(* IEC 61131-3 sources: plc-st-coding-agent/progress/evidence/f14_v10_full_20261113/jobs/codex_minimax-m27 (part 3) *)

(* ---- public-hard-05.candidate_02.st ---- *)
FUNCTION_BLOCK ArmController
VAR_INPUT
    ManualMode : BOOL;
    SingleStepMode : BOOL;
    SingleCycleMode : BOOL;
    ContinuousMode : BOOL;
    EmergencyStop : BOOL;
    Start : BOOL;
    DownButton : BOOL;
    UpButton : BOOL;
    LeftButton : BOOL;
    RightButton : BOOL;
    GripButton : BOOL;
    ReleaseButton : BOOL;
    DownLimitSwitch : BOOL;
    UpLimitSwitch : BOOL;
    LeftLimitSwitch : BOOL;
    RightLimitSwitch : BOOL;
    GripLimitSwitch : BOOL;
    ReleaseLimitSwitch : BOOL;
END_VAR
VAR_OUTPUT
    MoveDown : BOOL := FALSE;
    MoveUp : BOOL := FALSE;
    MoveLeft : BOOL := FALSE;
    MoveRight : BOOL := FALSE;
    ActivateGrip : BOOL := FALSE;
    ActivateRelease : BOOL := FALSE;
END_VAR
VAR
    step : INT := 0;
    startRisingEdge : R_TRIG;
    running : BOOL := FALSE;
    cycleComplete : BOOL := FALSE;
END_VAR

(* ENGINEERING_CONTRACT
| Output/State      | Activation       | Retention       | Reset/Deactivation             | Same-Scan Priority    | Units/Boundaries      |
|-------------------|------------------|-----------------|---------------------------------|-----------------------|-----------------------|
| MoveDown/Up/Left/Right | Edge/start/trig | Hold until done | EmergencyStop(FALSE), mode end  | Output latches stop   | BOOL, limit-based     |
| ActivateGrip/Release   | Edge/start/trig | Hold until done | EmergencyStop(FALSE), mode end  | Output latches stop   | BOOL, limit-based     |
| step[0..8]        | Start rising edge| Retained        | EmergencyStop(FALSE), mode end  | Initialized to 0      | INT, wrap to 0 at 8   |
| running           | Start rising edge| Retained        | EmergencyStop(FALSE), cycle end | FALSE when E-Stop     | BOOL, auto in cycle   |
| cycleComplete     | step=8 & done    | Retained        | Start rising edge               | Set only once         | BOOL, latched         |

PUB clause coverage:
- PUB001: Manual mode direct button control with limit checking
- PUB002-PUB007: Single step sequence (8 steps, Start advances)
- PUB008-PUB011: Single cycle executes full sequence once
- PUB012-PUB015: Continuous mode repeats cycle
- PUB016-PUB018: Emergency stop (FALSE=triggered) stops all outputs
- PUB019-PUB020: Grip/Release limit switches for completion feedback

Behavior:
- EmergencyStop=FALSE: All outputs=0, running=FALSE, step NOT reset (resume capability)
- Initial state: step=0, running=FALSE, all outputs=FALSE
- Caller ensures mutually exclusive mode inputs
*)
(* CONTRACT_RULES [] *)

startRisingEdge(CLK := Start);
running := running OR (startRisingEdge.Q AND (SingleStepMode OR SingleCycleMode OR ContinuousMode));

IF EmergencyStop = FALSE THEN
    MoveDown := FALSE;
    MoveUp := FALSE;
    MoveLeft := FALSE;
    MoveRight := FALSE;
    ActivateGrip := FALSE;
    ActivateRelease := FALSE;
    running := FALSE;
    cycleComplete := FALSE;
ELSE
    IF ManualMode THEN
        step := 0;
        running := FALSE;

        IF DownButton AND NOT DownLimitSwitch THEN
            MoveDown := TRUE;
        ELSIF UpButton AND NOT UpLimitSwitch THEN
            MoveUp := TRUE;
        ELSIF LeftButton AND NOT LeftLimitSwitch THEN
            MoveLeft := TRUE;
        ELSIF RightButton AND NOT RightLimitSwitch THEN
            MoveRight := TRUE;
        END_IF;

        IF GripButton THEN
            ActivateGrip := TRUE;
        END_IF;
        IF ReleaseButton THEN
            ActivateRelease := TRUE;
        END_IF;

    ELSIF SingleStepMode THEN
        IF startRisingEdge.Q AND NOT running THEN
            running := TRUE;
        END_IF;

        IF running THEN
            CASE step OF
                0:
                    IF UpLimitSwitch THEN
                        MoveDown := TRUE;
                        IF DownLimitSwitch THEN
                            MoveDown := FALSE;
                            step := 1;
                        END_IF;
                    END_IF;
                1:
                    MoveDown := FALSE;
                    ActivateGrip := TRUE;
                    IF GripLimitSwitch THEN
                        ActivateGrip := FALSE;
                        step := 2;
                    END_IF;
                2:
                    ActivateGrip := FALSE;
                    MoveUp := TRUE;
                    IF UpLimitSwitch THEN
                        MoveUp := FALSE;
                        step := 3;
                    END_IF;
                3:
                    MoveUp := FALSE;
                    MoveRight := TRUE;
                    IF RightLimitSwitch THEN
                        MoveRight := FALSE;
                        step := 4;
                    END_IF;
                4:
                    MoveRight := FALSE;
                    MoveDown := TRUE;
                    IF DownLimitSwitch THEN
                        MoveDown := FALSE;
                        step := 5;
                    END_IF;
                5:
                    MoveDown := FALSE;
                    ActivateRelease := TRUE;
                    IF ReleaseLimitSwitch THEN
                        ActivateRelease := FALSE;
                        step := 6;
                    END_IF;
                6:
                    ActivateRelease := FALSE;
                    MoveUp := TRUE;
                    IF UpLimitSwitch THEN
                        MoveUp := FALSE;
                        step := 7;
                    END_IF;
                7:
                    MoveUp := FALSE;
                    MoveLeft := TRUE;
                    IF LeftLimitSwitch THEN
                        MoveLeft := FALSE;
                        step := 8;
                    END_IF;
                8:
                    MoveLeft := FALSE;
                    running := FALSE;
                    step := 0;
            END_CASE;
        END_IF;

    ELSIF SingleCycleMode THEN
        IF startRisingEdge.Q AND NOT running AND NOT cycleComplete THEN
            running := TRUE;
        END_IF;

        IF running AND NOT cycleComplete THEN
            CASE step OF
                0:
                    IF UpLimitSwitch THEN
                        MoveDown := TRUE;
                        IF DownLimitSwitch THEN
                            MoveDown := FALSE;
                            step := 1;
                        END_IF;
                    END_IF;
                1:
                    MoveDown := FALSE;
                    ActivateGrip := TRUE;
                    IF GripLimitSwitch THEN
                        ActivateGrip := FALSE;
                        step := 2;
                    END_IF;
                2:
                    ActivateGrip := FALSE;
                    MoveUp := TRUE;
                    IF UpLimitSwitch THEN
                        MoveUp := FALSE;
                        step := 3;
                    END_IF;
                3:
                    MoveUp := FALSE;
                    MoveRight := TRUE;
                    IF RightLimitSwitch THEN
                        MoveRight := FALSE;
                        step := 4;
                    END_IF;
                4:
                    MoveRight := FALSE;
                    MoveDown := TRUE;
                    IF DownLimitSwitch THEN
                        MoveDown := FALSE;
                        step := 5;
                    END_IF;
                5:
                    MoveDown := FALSE;
                    ActivateRelease := TRUE;
                    IF ReleaseLimitSwitch THEN
                        ActivateRelease := FALSE;
                        step := 6;
                    END_IF;
                6:
                    ActivateRelease := FALSE;
                    MoveUp := TRUE;
                    IF UpLimitSwitch THEN
                        MoveUp := FALSE;
                        step := 7;
                    END_IF;
                7:
                    MoveUp := FALSE;
                    MoveLeft := TRUE;
                    IF LeftLimitSwitch THEN
                        MoveLeft := FALSE;
                        step := 8;
                    END_IF;
                8:
                    MoveLeft := FALSE;
                    running := FALSE;
                    cycleComplete := TRUE;
                    step := 0;
            END_CASE;
        END_IF;

    ELSIF ContinuousMode THEN
        IF startRisingEdge.Q AND NOT running THEN
            running := TRUE;
        END_IF;

        IF running THEN
            CASE step OF
                0:
                    IF UpLimitSwitch THEN
                        MoveDown := TRUE;
                        IF DownLimitSwitch THEN
                            MoveDown := FALSE;
                            step := 1;
                        END_IF;
                    END_IF;
                1:
                    MoveDown := FALSE;
                    ActivateGrip := TRUE;
                    IF GripLimitSwitch THEN
                        ActivateGrip := FALSE;
                        step := 2;
                    END_IF;
                2:
                    ActivateGrip := FALSE;
                    MoveUp := TRUE;
                    IF UpLimitSwitch THEN
                        MoveUp := FALSE;
                        step := 3;
                    END_IF;
                3:
                    MoveUp := FALSE;
                    MoveRight := TRUE;
                    IF RightLimitSwitch THEN
                        MoveRight := FALSE;
                        step := 4;
                    END_IF;
                4:
                    MoveRight := FALSE;
                    MoveDown := TRUE;
                    IF DownLimitSwitch THEN
                        MoveDown := FALSE;
                        step := 5;
                    END_IF;
                5:
                    MoveDown := FALSE;
                    ActivateRelease := TRUE;
                    IF ReleaseLimitSwitch THEN
                        ActivateRelease := FALSE;
                        step := 6;
                    END_IF;
                6:
                    ActivateRelease := FALSE;
                    MoveUp := TRUE;
                    IF UpLimitSwitch THEN
                        MoveUp := FALSE;
                        step := 7;
                    END_IF;
                7:
                    MoveUp := FALSE;
                    MoveLeft := TRUE;
                    IF LeftLimitSwitch THEN
                        MoveLeft := FALSE;
                        step := 0;
                    END_IF;
            END_CASE;
        END_IF;
    END_IF;
END_IF;

END_FUNCTION_BLOCK

(* ---- public-hard-05.candidate_03.st ---- *)
FUNCTION_BLOCK ArmController
VAR_INPUT
    ManualMode : BOOL;
    SingleStepMode : BOOL;
    SingleCycleMode : BOOL;
    ContinuousMode : BOOL;
    EmergencyStop : BOOL;
    Start : BOOL;
    DownButton : BOOL;
    UpButton : BOOL;
    LeftButton : BOOL;
    RightButton : BOOL;
    GripButton : BOOL;
    ReleaseButton : BOOL;
    DownLimitSwitch : BOOL;
    UpLimitSwitch : BOOL;
    LeftLimitSwitch : BOOL;
    RightLimitSwitch : BOOL;
    GripLimitSwitch : BOOL;
    ReleaseLimitSwitch : BOOL;
END_VAR
VAR_OUTPUT
    MoveDown : BOOL := FALSE;
    MoveUp : BOOL := FALSE;
    MoveLeft : BOOL := FALSE;
    MoveRight : BOOL := FALSE;
    ActivateGrip : BOOL := FALSE;
    ActivateRelease : BOOL := FALSE;
END_VAR
VAR
    step : INT := 0;
    startRisingEdge : R_TRIG;
    running : BOOL := FALSE;
    cycleComplete : BOOL := FALSE;
END_VAR

(* ENGINEERING_CONTRACT
| Output/State      | Activation       | Retention       | Reset/Deactivation             | Same-Scan Priority    | Units/Boundaries      |
|-------------------|------------------|-----------------|---------------------------------|-----------------------|-----------------------|
| MoveDown/Up/Left/Right | Edge/start/trig | Hold until done | EmergencyStop(FALSE), mode end  | Output latches stop   | BOOL, limit-based     |
| ActivateGrip/Release   | Edge/start/trig | Hold until done | EmergencyStop(FALSE), mode end  | Output latches stop   | BOOL, limit-based     |
| step[0..8]        | Start rising edge| Retained        | EmergencyStop(FALSE), mode end  | Initialized to 0      | INT, wrap to 0 at 8   |
| running           | Start rising edge| Retained        | EmergencyStop(FALSE), cycle end | FALSE when E-Stop     | BOOL, auto in cycle   |
| cycleComplete     | step=8 & done    | Retained        | Start rising edge               | Set only once         | BOOL, latched         |

PUB clause coverage:
- PUB001: Manual mode direct button control with limit checking
- PUB002-PUB007: Single step sequence (8 steps, Start advances)
- PUB008-PUB011: Single cycle executes full sequence once
- PUB012-PUB015: Continuous mode repeats cycle
- PUB016-PUB018: Emergency stop (FALSE=triggered) stops all outputs
- PUB019-PUB020: Grip/Release limit switches for completion feedback

Behavior:
- EmergencyStop=FALSE: All outputs=0, running=FALSE, cycleComplete NOT reset (resume capability)
- Initial state: step=0, running=FALSE, all outputs=FALSE
- Caller ensures mutually exclusive mode inputs
*)
(* CONTRACT_RULES [] *)

startRisingEdge(CLK := Start);
running := running OR (startRisingEdge.Q AND (SingleStepMode OR SingleCycleMode OR ContinuousMode));

IF EmergencyStop = FALSE THEN
    MoveDown := FALSE;
    MoveUp := FALSE;
    MoveLeft := FALSE;
    MoveRight := FALSE;
    ActivateGrip := FALSE;
    ActivateRelease := FALSE;
    running := FALSE;
    cycleComplete := FALSE;
ELSE
    IF ManualMode THEN
        step := 0;
        running := FALSE;
        MoveDown := FALSE;
        MoveUp := FALSE;
        MoveLeft := FALSE;
        MoveRight := FALSE;
        ActivateGrip := FALSE;
        ActivateRelease := FALSE;

        IF DownButton AND NOT DownLimitSwitch THEN
            MoveDown := TRUE;
        ELSIF UpButton AND NOT UpLimitSwitch THEN
            MoveUp := TRUE;
        ELSIF LeftButton AND NOT LeftLimitSwitch THEN
            MoveLeft := TRUE;
        ELSIF RightButton AND NOT RightLimitSwitch THEN
            MoveRight := TRUE;
        END_IF;

        IF GripButton THEN
            ActivateGrip := TRUE;
        END_IF;
        IF ReleaseButton THEN
            ActivateRelease := TRUE;
        END_IF;

    ELSIF SingleStepMode THEN
        MoveDown := FALSE;
        MoveUp := FALSE;
        MoveLeft := FALSE;
        MoveRight := FALSE;
        ActivateGrip := FALSE;
        ActivateRelease := FALSE;

        IF startRisingEdge.Q AND NOT running THEN
            running := TRUE;
        END_IF;

        IF running THEN
            CASE step OF
                0:
                    MoveDown := TRUE;
                    IF DownLimitSwitch THEN
                        MoveDown := FALSE;
                        step := 1;
                        running := FALSE;
                    END_IF;
                1:
                    ActivateGrip := TRUE;
                    IF GripLimitSwitch THEN
                        ActivateGrip := FALSE;
                        step := 2;
                        running := FALSE;
                    END_IF;
                2:
                    MoveUp := TRUE;
                    IF UpLimitSwitch THEN
                        MoveUp := FALSE;
                        step := 3;
                        running := FALSE;
                    END_IF;
                3:
                    MoveRight := TRUE;
                    IF RightLimitSwitch THEN
                        MoveRight := FALSE;
                        step := 4;
                        running := FALSE;
                    END_IF;
                4:
                    MoveDown := TRUE;
                    IF DownLimitSwitch THEN
                        MoveDown := FALSE;
                        step := 5;
                        running := FALSE;
                    END_IF;
                5:
                    ActivateRelease := TRUE;
                    IF ReleaseLimitSwitch THEN
                        ActivateRelease := FALSE;
                        step := 6;
                        running := FALSE;
                    END_IF;
                6:
                    MoveUp := TRUE;
                    IF UpLimitSwitch THEN
                        MoveUp := FALSE;
                        step := 7;
                        running := FALSE;
                    END_IF;
                7:
                    MoveLeft := TRUE;
                    IF LeftLimitSwitch THEN
                        MoveLeft := FALSE;
                        step := 8;
                        running := FALSE;
                    END_IF;
                8:
                    step := 0;
                    running := FALSE;
            END_CASE;
        END_IF;

    ELSIF SingleCycleMode THEN
        MoveDown := FALSE;
        MoveUp := FALSE;
        MoveLeft := FALSE;
        MoveRight := FALSE;
        ActivateGrip := FALSE;
        ActivateRelease := FALSE;

        IF startRisingEdge.Q AND NOT running AND NOT cycleComplete THEN
            running := TRUE;
        END_IF;

        IF running AND NOT cycleComplete THEN
            CASE step OF
                0:
                    MoveDown := TRUE;
                    IF DownLimitSwitch THEN
                        MoveDown := FALSE;
                        step := 1;
                    END_IF;
                1:
                    ActivateGrip := TRUE;
                    IF GripLimitSwitch THEN
                        ActivateGrip := FALSE;
                        step := 2;
                    END_IF;
                2:
                    MoveUp := TRUE;
                    IF UpLimitSwitch THEN
                        MoveUp := FALSE;
                        step := 3;
                    END_IF;
                3:
                    MoveRight := TRUE;
                    IF RightLimitSwitch THEN
                        MoveRight := FALSE;
                        step := 4;
                    END_IF;
                4:
                    MoveDown := TRUE;
                    IF DownLimitSwitch THEN
                        MoveDown := FALSE;
                        step := 5;
                    END_IF;
                5:
                    ActivateRelease := TRUE;
                    IF ReleaseLimitSwitch THEN
                        ActivateRelease := FALSE;
                        step := 6;
                    END_IF;
                6:
                    MoveUp := TRUE;
                    IF UpLimitSwitch THEN
                        MoveUp := FALSE;
                        step := 7;
                    END_IF;
                7:
                    MoveLeft := TRUE;
                    IF LeftLimitSwitch THEN
                        MoveLeft := FALSE;
                        step := 8;
                    END_IF;
                8:
                    MoveLeft := FALSE;
                    running := FALSE;
                    cycleComplete := TRUE;
                    step := 0;
            END_CASE;
        END_IF;

    ELSIF ContinuousMode THEN
        MoveDown := FALSE;
        MoveUp := FALSE;
        MoveLeft := FALSE;
        MoveRight := FALSE;
        ActivateGrip := FALSE;
        ActivateRelease := FALSE;

        IF startRisingEdge.Q AND NOT running THEN
            running := TRUE;
        END_IF;

        IF running THEN
            CASE step OF
                0:
                    MoveDown := TRUE;
                    IF DownLimitSwitch THEN
                        MoveDown := FALSE;
                        step := 1;
                    END_IF;
                1:
                    ActivateGrip := TRUE;
                    IF GripLimitSwitch THEN
                        ActivateGrip := FALSE;
                        step := 2;
                    END_IF;
                2:
                    MoveUp := TRUE;
                    IF UpLimitSwitch THEN
                        MoveUp := FALSE;
                        step := 3;
                    END_IF;
                3:
                    MoveRight := TRUE;
                    IF RightLimitSwitch THEN
                        MoveRight := FALSE;
                        step := 4;
                    END_IF;
                4:
                    MoveDown := TRUE;
                    IF DownLimitSwitch THEN
                        MoveDown := FALSE;
                        step := 5;
                    END_IF;
                5:
                    ActivateRelease := TRUE;
                    IF ReleaseLimitSwitch THEN
                        ActivateRelease := FALSE;
                        step := 6;
                    END_IF;
                6:
                    MoveUp := TRUE;
                    IF UpLimitSwitch THEN
                        MoveUp := FALSE;
                        step := 7;
                    END_IF;
                7:
                    MoveLeft := TRUE;
                    IF LeftLimitSwitch THEN
                        MoveLeft := FALSE;
                        step := 0;
                    END_IF;
            END_CASE;
        END_IF;
    END_IF;
END_IF;

END_FUNCTION_BLOCK

(* ---- public-hard-05.candidate_04.st ---- *)
FUNCTION_BLOCK ArmController
VAR_INPUT
    ManualMode : BOOL;
    SingleStepMode : BOOL;
    SingleCycleMode : BOOL;
    ContinuousMode : BOOL;
    EmergencyStop : BOOL;
    Start : BOOL;
    DownButton : BOOL;
    UpButton : BOOL;
    LeftButton : BOOL;
    RightButton : BOOL;
    GripButton : BOOL;
    ReleaseButton : BOOL;
    DownLimitSwitch : BOOL;
    UpLimitSwitch : BOOL;
    LeftLimitSwitch : BOOL;
    RightLimitSwitch : BOOL;
    GripLimitSwitch : BOOL;
    ReleaseLimitSwitch : BOOL;
END_VAR
VAR_OUTPUT
    MoveDown : BOOL := FALSE;
    MoveUp : BOOL := FALSE;
    MoveLeft : BOOL := FALSE;
    MoveRight : BOOL := FALSE;
    ActivateGrip : BOOL := FALSE;
    ActivateRelease : BOOL := FALSE;
END_VAR
VAR
    step : INT := 0;
    startRisingEdge : R_TRIG;
    running : BOOL := FALSE;
    cycleComplete : BOOL := FALSE;
END_VAR

(* ENGINEERING_CONTRACT
| Output/State      | Activation       | Retention       | Reset/Deactivation             | Same-Scan Priority    | Units/Boundaries      |
|-------------------|------------------|-----------------|---------------------------------|-----------------------|-----------------------|
| MoveDown/Up/Left/Right | Step-dependent | Hold until done | EmergencyStop(FALSE), mode end  | Output based on step  | BOOL, limit-based     |
| ActivateGrip/Release   | Step-dependent | Hold until done | EmergencyStop(FALSE), mode end  | Output based on step  | BOOL, limit-based     |
| step[0..7]        | Limit reached    | Retained        | EmergencyStop(FALSE), mode end  | Initialized to 0      | INT, wrap to 0 at 7   |
| running           | Start rising edge| Retained        | EmergencyStop(FALSE), cycle end | FALSE when E-Stop     | BOOL, auto in cycle   |
| cycleComplete     | step=7 & done    | Retained        | Start rising edge               | Set only once         | BOOL, latched         |

PUB clause coverage:
- PUB001: Manual mode direct button control with limit checking
- PUB002-PUB007: Single step sequence (8 steps, Start advances)
- PUB008-PUB011: Single cycle executes full sequence once
- PUB012-PUB015: Continuous mode repeats cycle
- PUB016-PUB018: Emergency stop (FALSE=triggered) stops all outputs
- PUB019-PUB020: Grip/Release limit switches for completion feedback

Behavior:
- EmergencyStop=FALSE: All outputs=0, running=FALSE, cycleComplete NOT reset
- Initial state: step=0, running=FALSE, all outputs=FALSE
- Step advances only when corresponding limit switch condition is met
- Outputs set based on current step, not after condition evaluation
*)
(* CONTRACT_RULES [] *)

startRisingEdge(CLK := Start);

IF EmergencyStop = FALSE THEN
    MoveDown := FALSE;
    MoveUp := FALSE;
    MoveLeft := FALSE;
    MoveRight := FALSE;
    ActivateGrip := FALSE;
    ActivateRelease := FALSE;
    running := FALSE;
    cycleComplete := FALSE;
    step := 0;
ELSE
    IF ManualMode THEN
        step := 0;
        running := FALSE;
        MoveDown := DownButton AND NOT DownLimitSwitch;
        MoveUp := UpButton AND NOT UpLimitSwitch;
        MoveLeft := LeftButton AND NOT LeftLimitSwitch;
        MoveRight := RightButton AND NOT RightLimitSwitch;
        ActivateGrip := GripButton;
        ActivateRelease := ReleaseButton;

    ELSIF SingleStepMode THEN
        MoveDown := FALSE;
        MoveUp := FALSE;
        MoveLeft := FALSE;
        MoveRight := FALSE;
        ActivateGrip := FALSE;
        ActivateRelease := FALSE;

        IF startRisingEdge.Q AND NOT running THEN
            running := TRUE;
        END_IF;

        IF running THEN
            CASE step OF
                0:
                    IF NOT DownLimitSwitch THEN
                        MoveDown := TRUE;
                    END_IF;
                    IF DownLimitSwitch THEN
                        step := 1;
                        running := FALSE;
                    END_IF;
                1:
                    IF NOT GripLimitSwitch THEN
                        ActivateGrip := TRUE;
                    END_IF;
                    IF GripLimitSwitch THEN
                        step := 2;
                        running := FALSE;
                    END_IF;
                2:
                    IF NOT UpLimitSwitch THEN
                        MoveUp := TRUE;
                    END_IF;
                    IF UpLimitSwitch THEN
                        step := 3;
                        running := FALSE;
                    END_IF;
                3:
                    IF NOT RightLimitSwitch THEN
                        MoveRight := TRUE;
                    END_IF;
                    IF RightLimitSwitch THEN
                        step := 4;
                        running := FALSE;
                    END_IF;
                4:
                    IF NOT DownLimitSwitch THEN
                        MoveDown := TRUE;
                    END_IF;
                    IF DownLimitSwitch THEN
                        step := 5;
                        running := FALSE;
                    END_IF;
                5:
                    IF NOT ReleaseLimitSwitch THEN
                        ActivateRelease := TRUE;
                    END_IF;
                    IF ReleaseLimitSwitch THEN
                        step := 6;
                        running := FALSE;
                    END_IF;
                6:
                    IF NOT UpLimitSwitch THEN
                        MoveUp := TRUE;
                    END_IF;
                    IF UpLimitSwitch THEN
                        step := 7;
                        running := FALSE;
                    END_IF;
                7:
                    IF NOT LeftLimitSwitch THEN
                        MoveLeft := TRUE;
                    END_IF;
                    IF LeftLimitSwitch THEN
                        step := 0;
                        running := FALSE;
                    END_IF;
            END_CASE;
        END_IF;

    ELSIF SingleCycleMode THEN
        MoveDown := FALSE;
        MoveUp := FALSE;
        MoveLeft := FALSE;
        MoveRight := FALSE;
        ActivateGrip := FALSE;
        ActivateRelease := FALSE;

        IF startRisingEdge.Q AND NOT running AND NOT cycleComplete THEN
            running := TRUE;
        END_IF;

        IF running THEN
            CASE step OF
                0:
                    IF NOT DownLimitSwitch THEN
                        MoveDown := TRUE;
                    END_IF;
                    IF DownLimitSwitch THEN
                        step := 1;
                    END_IF;
                1:
                    IF NOT GripLimitSwitch THEN
                        ActivateGrip := TRUE;
                    END_IF;
                    IF GripLimitSwitch THEN
                        step := 2;
                    END_IF;
                2:
                    IF NOT UpLimitSwitch THEN
                        MoveUp := TRUE;
                    END_IF;
                    IF UpLimitSwitch THEN
                        step := 3;
                    END_IF;
                3:
                    IF NOT RightLimitSwitch THEN
                        MoveRight := TRUE;
                    END_IF;
                    IF RightLimitSwitch THEN
                        step := 4;
                    END_IF;
                4:
                    IF NOT DownLimitSwitch THEN
                        MoveDown := TRUE;
                    END_IF;
                    IF DownLimitSwitch THEN
                        step := 5;
                    END_IF;
                5:
                    IF NOT ReleaseLimitSwitch THEN
                        ActivateRelease := TRUE;
                    END_IF;
                    IF ReleaseLimitSwitch THEN
                        step := 6;
                    END_IF;
                6:
                    IF NOT UpLimitSwitch THEN
                        MoveUp := TRUE;
                    END_IF;
                    IF UpLimitSwitch THEN
                        step := 7;
                    END_IF;
                7:
                    IF NOT LeftLimitSwitch THEN
                        MoveLeft := TRUE;
                    END_IF;
                    IF LeftLimitSwitch THEN
                        running := FALSE;
                        cycleComplete := TRUE;
                        step := 0;
                    END_IF;
            END_CASE;
        END_IF;

    ELSIF ContinuousMode THEN
        MoveDown := FALSE;
        MoveUp := FALSE;
        MoveLeft := FALSE;
        MoveRight := FALSE;
        ActivateGrip := FALSE;
        ActivateRelease := FALSE;

        IF startRisingEdge.Q AND NOT running THEN
            running := TRUE;
        END_IF;

        IF running THEN
            CASE step OF
                0:
                    IF NOT DownLimitSwitch THEN
                        MoveDown := TRUE;
                    END_IF;
                    IF DownLimitSwitch THEN
                        step := 1;
                    END_IF;
                1:
                    IF NOT GripLimitSwitch THEN
                        ActivateGrip := TRUE;
                    END_IF;
                    IF GripLimitSwitch THEN
                        step := 2;
                    END_IF;
                2:
                    IF NOT UpLimitSwitch THEN
                        MoveUp := TRUE;
                    END_IF;
                    IF UpLimitSwitch THEN
                        step := 3;
                    END_IF;
                3:
                    IF NOT RightLimitSwitch THEN
                        MoveRight := TRUE;
                    END_IF;
                    IF RightLimitSwitch THEN
                        step := 4;
                    END_IF;
                4:
                    IF NOT DownLimitSwitch THEN
                        MoveDown := TRUE;
                    END_IF;
                    IF DownLimitSwitch THEN
                        step := 5;
                    END_IF;
                5:
                    IF NOT ReleaseLimitSwitch THEN
                        ActivateRelease := TRUE;
                    END_IF;
                    IF ReleaseLimitSwitch THEN
                        step := 6;
                    END_IF;
                6:
                    IF NOT UpLimitSwitch THEN
                        MoveUp := TRUE;
                    END_IF;
                    IF UpLimitSwitch THEN
                        step := 7;
                    END_IF;
                7:
                    IF NOT LeftLimitSwitch THEN
                        MoveLeft := TRUE;
                    END_IF;
                    IF LeftLimitSwitch THEN
                        step := 0;
                    END_IF;
            END_CASE;
        END_IF;
    END_IF;
END_IF;

END_FUNCTION_BLOCK

(* ---- public-hard-05.raw_candidate_01.st ---- *)
FUNCTION_BLOCK ArmController
VAR_INPUT
    ManualMode : BOOL;
    SingleStepMode : BOOL;
    SingleCycleMode : BOOL;
    ContinuousMode : BOOL;
    EmergencyStop : BOOL;
    Start : BOOL;
    DownButton : BOOL;
    UpButton : BOOL;
    LeftButton : BOOL;
    RightButton : BOOL;
    GripButton : BOOL;
    ReleaseButton : BOOL;
    DownLimitSwitch : BOOL;
    UpLimitSwitch : BOOL;
    LeftLimitSwitch : BOOL;
    RightLimitSwitch : BOOL;
    GripLimitSwitch : BOOL;
    ReleaseLimitSwitch : BOOL;
END_VAR
VAR_OUTPUT
    MoveDown : BOOL := FALSE;
    MoveUp : BOOL := FALSE;
    MoveLeft : BOOL := FALSE;
    MoveRight : BOOL := FALSE;
    ActivateGrip : BOOL := FALSE;
    ActivateRelease : BOOL := FALSE;
END_VAR
VAR
    step : INT := 0;
    startRisingEdge : R_TRIG;
    running : BOOL := FALSE;
    cycleComplete : BOOL := FALSE;
    tmpRunning : BOOL;
END_VAR

(* ENGINEERING_CONTRACT
| Output/State      | Activation       | Retention       | Reset/Deactivation             | Same-Scan Priority    | Units/Boundaries      |
|-------------------|------------------|-----------------|---------------------------------|-----------------------|-----------------------|
| MoveDown/Up/Left/Right | Edge/start/trig | Hold until done | EmergencyStop(FALSE), mode end  | Output latches stop   | BOOL, limit-based     |
| ActivateGrip/Release   | Edge/start/trig | Hold until done | EmergencyStop(FALSE), mode end  | Output latches stop   | BOOL, limit-based     |
| step[0..8]        | Start rising edge| Retained        | EmergencyStop(FALSE), mode end  | Initialized to 0      | INT, wrap to 0 at 8   |
| running           | Start rising edge| Retained        | EmergencyStop(FALSE), cycle end | FALSE when E-Stop     | BOOL, auto in cycle   |
| cycleComplete     | step=8 & done    | Retained        | Start rising edge               | Set only once         | BOOL, latched         |

PUB clause coverage:
- PUB001: Manual mode direct button control with limit checking
- PUB002-PUB007: Single step sequence (8 steps, Start advances)
- PUB008-PUB011: Single cycle executes full sequence once
- PUB012-PUB015: Continuous mode repeats cycle
- PUB016-PUB018: Emergency stop (FALSE=triggered) stops all outputs
- PUB019-PUB020: Grip/Release limit switches for completion feedback

Behavior:
- EmergencyStop=FALSE: All outputs=0, running=FALSE, step NOT reset (resume capability)
- Initial state: step=0, running=FALSE, all outputs=FALSE
- Caller ensures mutually exclusive mode inputs
*)
(* CONTRACT_RULES [] *)

tmpRunning := running;

startRisingEdge(CLK := Start);
running := running OR (startRisingEdge.Q AND (SingleStepMode OR SingleCycleMode OR ContinuousMode));

IF EmergencyStop = FALSE THEN
    MoveDown := FALSE;
    MoveUp := FALSE;
    MoveLeft := FALSE;
    MoveRight := FALSE;
    ActivateGrip := FALSE;
    ActivateRelease := FALSE;
    running := FALSE;
    cycleComplete := FALSE;
ELSE
    IF ManualMode THEN
        step := 0;
        running := FALSE;

        IF DownButton AND NOT DownLimitSwitch THEN
            MoveDown := TRUE;
        END_IF
        IF UpButton AND NOT UpLimitSwitch THEN
            MoveUp := TRUE;
        END_IF
        IF LeftButton AND NOT LeftLimitSwitch THEN
            MoveLeft := TRUE;
        END_IF
        IF RightButton AND NOT RightLimitSwitch THEN
            MoveRight := TRUE;
        END_IF
        IF GripButton THEN
            ActivateGrip := TRUE;
        END_IF
        IF ReleaseButton THEN
            ActivateRelease := TRUE;
        END_IF

    ELSIF SingleStepMode THEN
        IF startRisingEdge.Q AND NOT running THEN
            running := TRUE;
        END_IF

        IF running THEN
            CASE step OF
                0:
                    IF UpLimitSwitch THEN
                        MoveDown := TRUE;
                        IF DownLimitSwitch THEN
                            MoveDown := FALSE;
                            step := 1;
                        END_IF
                    END_IF
                1:
                    MoveDown := FALSE;
                    ActivateGrip := TRUE;
                    IF GripLimitSwitch THEN
                        ActivateGrip := FALSE;
                        step := 2;
                    END_IF
                2:
                    ActivateGrip := FALSE;
                    MoveUp := TRUE;
                    IF UpLimitSwitch THEN
                        MoveUp := FALSE;
                        step := 3;
                    END_IF
                3:
                    MoveUp := FALSE;
                    MoveRight := TRUE;
                    IF RightLimitSwitch THEN
                        MoveRight := FALSE;
                        step := 4;
                    END_IF
                4:
                    MoveRight := FALSE;
                    MoveDown := TRUE;
                    IF DownLimitSwitch THEN
                        MoveDown := FALSE;
                        step := 5;
                    END_IF
                5:
                    MoveDown := FALSE;
                    ActivateRelease := TRUE;
                    IF ReleaseLimitSwitch THEN
                        ActivateRelease := FALSE;
                        step := 6;
                    END_IF
                6:
                    ActivateRelease := FALSE;
                    MoveUp := TRUE;
                    IF UpLimitSwitch THEN
                        MoveUp := FALSE;
                        step := 7;
                    END_IF
                7:
                    MoveUp := FALSE;
                    MoveLeft := TRUE;
                    IF LeftLimitSwitch THEN
                        MoveLeft := FALSE;
                        step := 8;
                    END_IF
                8:
                    MoveLeft := FALSE;
                    running := FALSE;
                    step := 0;
            END_CASE
        END_IF

    ELSIF SingleCycleMode THEN
        IF startRisingEdge.Q AND NOT running AND NOT cycleComplete THEN
            running := TRUE;
        END_IF

        IF running AND NOT cycleComplete THEN
            CASE step OF
                0:
                    IF UpLimitSwitch THEN
                        MoveDown := TRUE;
                        IF DownLimitSwitch THEN
                            MoveDown := FALSE;
                            step := 1;
                        END_IF
                    END_IF
                1:
                    MoveDown := FALSE;
                    ActivateGrip := TRUE;
                    IF GripLimitSwitch THEN
                        ActivateGrip := FALSE;
                        step := 2;
                    END_IF
                2:
                    ActivateGrip := FALSE;
                    MoveUp := TRUE;
                    IF UpLimitSwitch THEN
                        MoveUp := FALSE;
                        step := 3;
                    END_IF
                3:
                    MoveUp := FALSE;
                    MoveRight := TRUE;
                    IF RightLimitSwitch THEN
                        MoveRight := FALSE;
                        step := 4;
                    END_IF
                4:
                    MoveRight := FALSE;
                    MoveDown := TRUE;
                    IF DownLimitSwitch THEN
                        MoveDown := FALSE;
                        step := 5;
                    END_IF
                5:
                    MoveDown := FALSE;
                    ActivateRelease := TRUE;
                    IF ReleaseLimitSwitch THEN
                        ActivateRelease := FALSE;
                        step := 6;
                    END_IF
                6:
                    ActivateRelease := FALSE;
                    MoveUp := TRUE;
                    IF UpLimitSwitch THEN
                        MoveUp := FALSE;
                        step := 7;
                    END_IF
                7:
                    MoveUp := FALSE;
                    MoveLeft := TRUE;
                    IF LeftLimitSwitch THEN
                        MoveLeft := FALSE;
                        step := 8;
                    END_IF
                8:
                    MoveLeft := FALSE;
                    running := FALSE;
                    cycleComplete := TRUE;
                    step := 0;
            END_CASE
        END_IF

    ELSIF ContinuousMode THEN
        IF startRisingEdge.Q AND NOT running THEN
            running := TRUE;
        END_IF

        IF running THEN
            CASE step OF
                0:
                    IF UpLimitSwitch THEN
                        MoveDown := TRUE;
                        IF DownLimitSwitch THEN
                            MoveDown := FALSE;
                            step := 1;
                        END_IF
                    END_IF
                1:
                    MoveDown := FALSE;
                    ActivateGrip := TRUE;
                    IF GripLimitSwitch THEN
                        ActivateGrip := FALSE;
                        step := 2;
                    END_IF
                2:
                    ActivateGrip := FALSE;
                    MoveUp := TRUE;
                    IF UpLimitSwitch THEN
                        MoveUp := FALSE;
                        step := 3;
                    END_IF
                3:
                    MoveUp := FALSE;
                    MoveRight := TRUE;
                    IF RightLimitSwitch THEN
                        MoveRight := FALSE;
                        step := 4;
                    END_IF
                4:
                    MoveRight := FALSE;
                    MoveDown := TRUE;
                    IF DownLimitSwitch THEN
                        MoveDown := FALSE;
                        step := 5;
                    END_IF
                5:
                    MoveDown := FALSE;
                    ActivateRelease := TRUE;
                    IF ReleaseLimitSwitch THEN
                        ActivateRelease := FALSE;
                        step := 6;
                    END_IF
                6:
                    ActivateRelease := FALSE;
                    MoveUp := TRUE;
                    IF UpLimitSwitch THEN
                        MoveUp := FALSE;
                        step := 7;
                    END_IF
                7:
                    MoveUp := FALSE;
                    MoveLeft := TRUE;
                    IF LeftLimitSwitch THEN
                        MoveLeft := FALSE;
                        step := 0;
                    END_IF
            END_CASE
        END_IF
    END_IF
END_IF

END_FUNCTION_BLOCK

(* ---- public-hard-05.raw_candidate_02.st ---- *)
FUNCTION_BLOCK ArmController
VAR_INPUT
    ManualMode : BOOL;
    SingleStepMode : BOOL;
    SingleCycleMode : BOOL;
    ContinuousMode : BOOL;
    EmergencyStop : BOOL;
    Start : BOOL;
    DownButton : BOOL;
    UpButton : BOOL;
    LeftButton : BOOL;
    RightButton : BOOL;
    GripButton : BOOL;
    ReleaseButton : BOOL;
    DownLimitSwitch : BOOL;
    UpLimitSwitch : BOOL;
    LeftLimitSwitch : BOOL;
    RightLimitSwitch : BOOL;
    GripLimitSwitch : BOOL;
    ReleaseLimitSwitch : BOOL;
END_VAR
VAR_OUTPUT
    MoveDown : BOOL := FALSE;
    MoveUp : BOOL := FALSE;
    MoveLeft : BOOL := FALSE;
    MoveRight : BOOL := FALSE;
    ActivateGrip : BOOL := FALSE;
    ActivateRelease : BOOL := FALSE;
END_VAR
VAR
    step : INT := 0;
    startRisingEdge : R_TRIG;
    running : BOOL := FALSE;
    cycleComplete : BOOL := FALSE;
END_VAR

(* ENGINEERING_CONTRACT
| Output/State      | Activation       | Retention       | Reset/Deactivation             | Same-Scan Priority    | Units/Boundaries      |
|-------------------|------------------|-----------------|---------------------------------|-----------------------|-----------------------|
| MoveDown/Up/Left/Right | Edge/start/trig | Hold until done | EmergencyStop(FALSE), mode end  | Output latches stop   | BOOL, limit-based     |
| ActivateGrip/Release   | Edge/start/trig | Hold until done | EmergencyStop(FALSE), mode end  | Output latches stop   | BOOL, limit-based     |
| step[0..8]        | Start rising edge| Retained        | EmergencyStop(FALSE), mode end  | Initialized to 0      | INT, wrap to 0 at 8   |
| running           | Start rising edge| Retained        | EmergencyStop(FALSE), cycle end | FALSE when E-Stop     | BOOL, auto in cycle   |
| cycleComplete     | step=8 & done    | Retained        | Start rising edge               | Set only once         | BOOL, latched         |

PUB clause coverage:
- PUB001: Manual mode direct button control with limit checking
- PUB002-PUB007: Single step sequence (8 steps, Start advances)
- PUB008-PUB011: Single cycle executes full sequence once
- PUB012-PUB015: Continuous mode repeats cycle
- PUB016-PUB018: Emergency stop (FALSE=triggered) stops all outputs
- PUB019-PUB020: Grip/Release limit switches for completion feedback

Behavior:
- EmergencyStop=FALSE: All outputs=0, running=FALSE, step NOT reset (resume capability)
- Initial state: step=0, running=FALSE, all outputs=FALSE
- Caller ensures mutually exclusive mode inputs
*)
(* CONTRACT_RULES [] *)

startRisingEdge(CLK := Start);
running := running OR (startRisingEdge.Q AND (SingleStepMode OR SingleCycleMode OR ContinuousMode));

IF EmergencyStop = FALSE THEN
    MoveDown := FALSE;
    MoveUp := FALSE;
    MoveLeft := FALSE;
    MoveRight := FALSE;
    ActivateGrip := FALSE;
    ActivateRelease := FALSE;
    running := FALSE;
    cycleComplete := FALSE;
ELSE
    IF ManualMode THEN
        step := 0;
        running := FALSE;

        IF DownButton AND NOT DownLimitSwitch THEN
            MoveDown := TRUE;
        ELSIF UpButton AND NOT UpLimitSwitch THEN
            MoveUp := TRUE;
        ELSIF LeftButton AND NOT LeftLimitSwitch THEN
            MoveLeft := TRUE;
        ELSIF RightButton AND NOT RightLimitSwitch THEN
            MoveRight := TRUE;
        END_IF;

        IF GripButton THEN
            ActivateGrip := TRUE;
        END_IF;
        IF ReleaseButton THEN
            ActivateRelease := TRUE;
        END_IF;

    ELSIF SingleStepMode THEN
        IF startRisingEdge.Q AND NOT running THEN
            running := TRUE;
        END_IF;

        IF running THEN
            CASE step OF
                0:
                    IF UpLimitSwitch THEN
                        MoveDown := TRUE;
                        IF DownLimitSwitch THEN
                            MoveDown := FALSE;
                            step := 1;
                        END_IF;
                    END_IF;
                1:
                    MoveDown := FALSE;
                    ActivateGrip := TRUE;
                    IF GripLimitSwitch THEN
                        ActivateGrip := FALSE;
                        step := 2;
                    END_IF;
                2:
                    ActivateGrip := FALSE;
                    MoveUp := TRUE;
                    IF UpLimitSwitch THEN
                        MoveUp := FALSE;
                        step := 3;
                    END_IF;
                3:
                    MoveUp := FALSE;
                    MoveRight := TRUE;
                    IF RightLimitSwitch THEN
                        MoveRight := FALSE;
                        step := 4;
                    END_IF;
                4:
                    MoveRight := FALSE;
                    MoveDown := TRUE;
                    IF DownLimitSwitch THEN
                        MoveDown := FALSE;
                        step := 5;
                    END_IF;
                5:
                    MoveDown := FALSE;
                    ActivateRelease := TRUE;
                    IF ReleaseLimitSwitch THEN
                        ActivateRelease := FALSE;
                        step := 6;
                    END_IF;
                6:
                    ActivateRelease := FALSE;
                    MoveUp := TRUE;
                    IF UpLimitSwitch THEN
                        MoveUp := FALSE;
                        step := 7;
                    END_IF;
                7:
                    MoveUp := FALSE;
                    MoveLeft := TRUE;
                    IF LeftLimitSwitch THEN
                        MoveLeft := FALSE;
                        step := 8;
                    END_IF;
                8:
                    MoveLeft := FALSE;
                    running := FALSE;
                    step := 0;
            END_CASE;
        END_IF;

    ELSIF SingleCycleMode THEN
        IF startRisingEdge.Q AND NOT running AND NOT cycleComplete THEN
            running := TRUE;
        END_IF;

        IF running AND NOT cycleComplete THEN
            CASE step OF
                0:
                    IF UpLimitSwitch THEN
                        MoveDown := TRUE;
                        IF DownLimitSwitch THEN
                            MoveDown := FALSE;
                            step := 1;
                        END_IF;
                    END_IF;
                1:
                    MoveDown := FALSE;
                    ActivateGrip := TRUE;
                    IF GripLimitSwitch THEN
                        ActivateGrip := FALSE;
                        step := 2;
                    END_IF;
                2:
                    ActivateGrip := FALSE;
                    MoveUp := TRUE;
                    IF UpLimitSwitch THEN
                        MoveUp := FALSE;
                        step := 3;
                    END_IF;
                3:
                    MoveUp := FALSE;
                    MoveRight := TRUE;
                    IF RightLimitSwitch THEN
                        MoveRight := FALSE;
                        step := 4;
                    END_IF;
                4:
                    MoveRight := FALSE;
                    MoveDown := TRUE;
                    IF DownLimitSwitch THEN
                        MoveDown := FALSE;
                        step := 5;
                    END_IF;
                5:
                    MoveDown := FALSE;
                    ActivateRelease := TRUE;
                    IF ReleaseLimitSwitch THEN
                        ActivateRelease := FALSE;
                        step := 6;
                    END_IF;
                6:
                    ActivateRelease := FALSE;
                    MoveUp := TRUE;
                    IF UpLimitSwitch THEN
                        MoveUp := FALSE;
                        step := 7;
                    END_IF;
                7:
                    MoveUp := FALSE;
                    MoveLeft := TRUE;
                    IF LeftLimitSwitch THEN
                        MoveLeft := FALSE;
                        step := 8;
                    END_IF;
                8:
                    MoveLeft := FALSE;
                    running := FALSE;
                    cycleComplete := TRUE;
                    step := 0;
            END_CASE;
        END_IF;

    ELSIF ContinuousMode THEN
        IF startRisingEdge.Q AND NOT running THEN
            running := TRUE;
        END_IF;

        IF running THEN
            CASE step OF
                0:
                    IF UpLimitSwitch THEN
                        MoveDown := TRUE;
                        IF DownLimitSwitch THEN
                            MoveDown := FALSE;
                            step := 1;
                        END_IF;
                    END_IF;
                1:
                    MoveDown := FALSE;
                    ActivateGrip := TRUE;
                    IF GripLimitSwitch THEN
                        ActivateGrip := FALSE;
                        step := 2;
                    END_IF;
                2:
                    ActivateGrip := FALSE;
                    MoveUp := TRUE;
                    IF UpLimitSwitch THEN
                        MoveUp := FALSE;
                        step := 3;
                    END_IF;
                3:
                    MoveUp := FALSE;
                    MoveRight := TRUE;
                    IF RightLimitSwitch THEN
                        MoveRight := FALSE;
                        step := 4;
                    END_IF;
                4:
                    MoveRight := FALSE;
                    MoveDown := TRUE;
                    IF DownLimitSwitch THEN
                        MoveDown := FALSE;
                        step := 5;
                    END_IF;
                5:
                    MoveDown := FALSE;
                    ActivateRelease := TRUE;
                    IF ReleaseLimitSwitch THEN
                        ActivateRelease := FALSE;
                        step := 6;
                    END_IF;
                6:
                    ActivateRelease := FALSE;
                    MoveUp := TRUE;
                    IF UpLimitSwitch THEN
                        MoveUp := FALSE;
                        step := 7;
                    END_IF;
                7:
                    MoveUp := FALSE;
                    MoveLeft := TRUE;
                    IF LeftLimitSwitch THEN
                        MoveLeft := FALSE;
                        step := 0;
                    END_IF;
            END_CASE;
        END_IF;
    END_IF;
END_IF;

END_FUNCTION_BLOCK

(* ---- public-hard-05.raw_candidate_03.st ---- *)
FUNCTION_BLOCK ArmController
VAR_INPUT
    ManualMode : BOOL;
    SingleStepMode : BOOL;
    SingleCycleMode : BOOL;
    ContinuousMode : BOOL;
    EmergencyStop : BOOL;
    Start : BOOL;
    DownButton : BOOL;
    UpButton : BOOL;
    LeftButton : BOOL;
    RightButton : BOOL;
    GripButton : BOOL;
    ReleaseButton : BOOL;
    DownLimitSwitch : BOOL;
    UpLimitSwitch : BOOL;
    LeftLimitSwitch : BOOL;
    RightLimitSwitch : BOOL;
    GripLimitSwitch : BOOL;
    ReleaseLimitSwitch : BOOL;
END_VAR
VAR_OUTPUT
    MoveDown : BOOL := FALSE;
    MoveUp : BOOL := FALSE;
    MoveLeft : BOOL := FALSE;
    MoveRight : BOOL := FALSE;
    ActivateGrip : BOOL := FALSE;
    ActivateRelease : BOOL := FALSE;
END_VAR
VAR
    step : INT := 0;
    startRisingEdge : R_TRIG;
    running : BOOL := FALSE;
    cycleComplete : BOOL := FALSE;
END_VAR

(* ENGINEERING_CONTRACT
| Output/State      | Activation       | Retention       | Reset/Deactivation             | Same-Scan Priority    | Units/Boundaries      |
|-------------------|------------------|-----------------|---------------------------------|-----------------------|-----------------------|
| MoveDown/Up/Left/Right | Edge/start/trig | Hold until done | EmergencyStop(FALSE), mode end  | Output latches stop   | BOOL, limit-based     |
| ActivateGrip/Release   | Edge/start/trig | Hold until done | EmergencyStop(FALSE), mode end  | Output latches stop   | BOOL, limit-based     |
| step[0..8]        | Start rising edge| Retained        | EmergencyStop(FALSE), mode end  | Initialized to 0      | INT, wrap to 0 at 8   |
| running           | Start rising edge| Retained        | EmergencyStop(FALSE), cycle end | FALSE when E-Stop     | BOOL, auto in cycle   |
| cycleComplete     | step=8 & done    | Retained        | Start rising edge               | Set only once         | BOOL, latched         |

PUB clause coverage:
- PUB001: Manual mode direct button control with limit checking
- PUB002-PUB007: Single step sequence (8 steps, Start advances)
- PUB008-PUB011: Single cycle executes full sequence once
- PUB012-PUB015: Continuous mode repeats cycle
- PUB016-PUB018: Emergency stop (FALSE=triggered) stops all outputs
- PUB019-PUB020: Grip/Release limit switches for completion feedback

Behavior:
- EmergencyStop=FALSE: All outputs=0, running=FALSE, cycleComplete NOT reset (resume capability)
- Initial state: step=0, running=FALSE, all outputs=FALSE
- Caller ensures mutually exclusive mode inputs
*)
(* CONTRACT_RULES [] *)

startRisingEdge(CLK := Start);
running := running OR (startRisingEdge.Q AND (SingleStepMode OR SingleCycleMode OR ContinuousMode));

IF EmergencyStop = FALSE THEN
    MoveDown := FALSE;
    MoveUp := FALSE;
    MoveLeft := FALSE;
    MoveRight := FALSE;
    ActivateGrip := FALSE;
    ActivateRelease := FALSE;
    running := FALSE;
    cycleComplete := FALSE;
ELSE
    IF ManualMode THEN
        step := 0;
        running := FALSE;
        MoveDown := FALSE;
        MoveUp := FALSE;
        MoveLeft := FALSE;
        MoveRight := FALSE;
        ActivateGrip := FALSE;
        ActivateRelease := FALSE;

        IF DownButton AND NOT DownLimitSwitch THEN
            MoveDown := TRUE;
        ELSIF UpButton AND NOT UpLimitSwitch THEN
            MoveUp := TRUE;
        ELSIF LeftButton AND NOT LeftLimitSwitch THEN
            MoveLeft := TRUE;
        ELSIF RightButton AND NOT RightLimitSwitch THEN
            MoveRight := TRUE;
        END_IF;

        IF GripButton THEN
            ActivateGrip := TRUE;
        END_IF;
        IF ReleaseButton THEN
            ActivateRelease := TRUE;
        END_IF;

    ELSIF SingleStepMode THEN
        MoveDown := FALSE;
        MoveUp := FALSE;
        MoveLeft := FALSE;
        MoveRight := FALSE;
        ActivateGrip := FALSE;
        ActivateRelease := FALSE;

        IF startRisingEdge.Q AND NOT running THEN
            running := TRUE;
        END_IF;

        IF running THEN
            CASE step OF
                0:
                    MoveDown := TRUE;
                    IF DownLimitSwitch THEN
                        MoveDown := FALSE;
                        step := 1;
                        running := FALSE;
                    END_IF;
                1:
                    ActivateGrip := TRUE;
                    IF GripLimitSwitch THEN
                        ActivateGrip := FALSE;
                        step := 2;
                        running := FALSE;
                    END_IF;
                2:
                    MoveUp := TRUE;
                    IF UpLimitSwitch THEN
                        MoveUp := FALSE;
                        step := 3;
                        running := FALSE;
                    END_IF;
                3:
                    MoveRight := TRUE;
                    IF RightLimitSwitch THEN
                        MoveRight := FALSE;
                        step := 4;
                        running := FALSE;
                    END_IF;
                4:
                    MoveDown := TRUE;
                    IF DownLimitSwitch THEN
                        MoveDown := FALSE;
                        step := 5;
                        running := FALSE;
                    END_IF;
                5:
                    ActivateRelease := TRUE;
                    IF ReleaseLimitSwitch THEN
                        ActivateRelease := FALSE;
                        step := 6;
                        running := FALSE;
                    END_IF;
                6:
                    MoveUp := TRUE;
                    IF UpLimitSwitch THEN
                        MoveUp := FALSE;
                        step := 7;
                        running := FALSE;
                    END_IF;
                7:
                    MoveLeft := TRUE;
                    IF LeftLimitSwitch THEN
                        MoveLeft := FALSE;
                        step := 8;
                        running := FALSE;
                    END_IF;
                8:
                    step := 0;
                    running := FALSE;
            END_CASE;
        END_IF;

    ELSIF SingleCycleMode THEN
        MoveDown := FALSE;
        MoveUp := FALSE;
        MoveLeft := FALSE;
        MoveRight := FALSE;
        ActivateGrip := FALSE;
        ActivateRelease := FALSE;

        IF startRisingEdge.Q AND NOT running AND NOT cycleComplete THEN
            running := TRUE;
        END_IF;

        IF running AND NOT cycleComplete THEN
            CASE step OF
                0:
                    MoveDown := TRUE;
                    IF DownLimitSwitch THEN
                        MoveDown := FALSE;
                        step := 1;
                    END_IF;
                1:
                    ActivateGrip := TRUE;
                    IF GripLimitSwitch THEN
                        ActivateGrip := FALSE;
                        step := 2;
                    END_IF;
                2:
                    MoveUp := TRUE;
                    IF UpLimitSwitch THEN
                        MoveUp := FALSE;
                        step := 3;
                    END_IF;
                3:
                    MoveRight := TRUE;
                    IF RightLimitSwitch THEN
                        MoveRight := FALSE;
                        step := 4;
                    END_IF;
                4:
                    MoveDown := TRUE;
                    IF DownLimitSwitch THEN
                        MoveDown := FALSE;
                        step := 5;
                    END_IF;
                5:
                    ActivateRelease := TRUE;
                    IF ReleaseLimitSwitch THEN
                        ActivateRelease := FALSE;
                        step := 6;
                    END_IF;
                6:
                    MoveUp := TRUE;
                    IF UpLimitSwitch THEN
                        MoveUp := FALSE;
                        step := 7;
                    END_IF;
                7:
                    MoveLeft := TRUE;
                    IF LeftLimitSwitch THEN
                        MoveLeft := FALSE;
                        step := 8;
                    END_IF;
                8:
                    MoveLeft := FALSE;
                    running := FALSE;
                    cycleComplete := TRUE;
                    step := 0;
            END_CASE;
        END_IF;

    ELSIF ContinuousMode THEN
        MoveDown := FALSE;
        MoveUp := FALSE;
        MoveLeft := FALSE;
        MoveRight := FALSE;
        ActivateGrip := FALSE;
        ActivateRelease := FALSE;

        IF startRisingEdge.Q AND NOT running THEN
            running := TRUE;
        END_IF;

        IF running THEN
            CASE step OF
                0:
                    MoveDown := TRUE;
                    IF DownLimitSwitch THEN
                        MoveDown := FALSE;
                        step := 1;
                    END_IF;
                1:
                    ActivateGrip := TRUE;
                    IF GripLimitSwitch THEN
                        ActivateGrip := FALSE;
                        step := 2;
                    END_IF;
                2:
                    MoveUp := TRUE;
                    IF UpLimitSwitch THEN
                        MoveUp := FALSE;
                        step := 3;
                    END_IF;
                3:
                    MoveRight := TRUE;
                    IF RightLimitSwitch THEN
                        MoveRight := FALSE;
                        step := 4;
                    END_IF;
                4:
                    MoveDown := TRUE;
                    IF DownLimitSwitch THEN
                        MoveDown := FALSE;
                        step := 5;
                    END_IF;
                5:
                    ActivateRelease := TRUE;
                    IF ReleaseLimitSwitch THEN
                        ActivateRelease := FALSE;
                        step := 6;
                    END_IF;
                6:
                    MoveUp := TRUE;
                    IF UpLimitSwitch THEN
                        MoveUp := FALSE;
                        step := 7;
                    END_IF;
                7:
                    MoveLeft := TRUE;
                    IF LeftLimitSwitch THEN
                        MoveLeft := FALSE;
                        step := 0;
                    END_IF;
            END_CASE;
        END_IF;
    END_IF;
END_IF;

END_FUNCTION_BLOCK

(* ---- public-hard-05.raw_candidate_04.st ---- *)
FUNCTION_BLOCK ArmController
VAR_INPUT
    ManualMode : BOOL;
    SingleStepMode : BOOL;
    SingleCycleMode : BOOL;
    ContinuousMode : BOOL;
    EmergencyStop : BOOL;
    Start : BOOL;
    DownButton : BOOL;
    UpButton : BOOL;
    LeftButton : BOOL;
    RightButton : BOOL;
    GripButton : BOOL;
    ReleaseButton : BOOL;
    DownLimitSwitch : BOOL;
    UpLimitSwitch : BOOL;
    LeftLimitSwitch : BOOL;
    RightLimitSwitch : BOOL;
    GripLimitSwitch : BOOL;
    ReleaseLimitSwitch : BOOL;
END_VAR
VAR_OUTPUT
    MoveDown : BOOL := FALSE;
    MoveUp : BOOL := FALSE;
    MoveLeft : BOOL := FALSE;
    MoveRight : BOOL := FALSE;
    ActivateGrip : BOOL := FALSE;
    ActivateRelease : BOOL := FALSE;
END_VAR
VAR
    step : INT := 0;
    startRisingEdge : R_TRIG;
    running : BOOL := FALSE;
    cycleComplete : BOOL := FALSE;
END_VAR

(* ENGINEERING_CONTRACT
| Output/State      | Activation       | Retention       | Reset/Deactivation             | Same-Scan Priority    | Units/Boundaries      |
|-------------------|------------------|-----------------|---------------------------------|-----------------------|-----------------------|
| MoveDown/Up/Left/Right | Step-dependent | Hold until done | EmergencyStop(FALSE), mode end  | Output based on step  | BOOL, limit-based     |
| ActivateGrip/Release   | Step-dependent | Hold until done | EmergencyStop(FALSE), mode end  | Output based on step  | BOOL, limit-based     |
| step[0..7]        | Limit reached    | Retained        | EmergencyStop(FALSE), mode end  | Initialized to 0      | INT, wrap to 0 at 7   |
| running           | Start rising edge| Retained        | EmergencyStop(FALSE), cycle end | FALSE when E-Stop     | BOOL, auto in cycle   |
| cycleComplete     | step=7 & done    | Retained        | Start rising edge               | Set only once         | BOOL, latched         |

PUB clause coverage:
- PUB001: Manual mode direct button control with limit checking
- PUB002-PUB007: Single step sequence (8 steps, Start advances)
- PUB008-PUB011: Single cycle executes full sequence once
- PUB012-PUB015: Continuous mode repeats cycle
- PUB016-PUB018: Emergency stop (FALSE=triggered) stops all outputs
- PUB019-PUB020: Grip/Release limit switches for completion feedback

Behavior:
- EmergencyStop=FALSE: All outputs=0, running=FALSE, cycleComplete NOT reset
- Initial state: step=0, running=FALSE, all outputs=FALSE
- Step advances only when corresponding limit switch condition is met
- Outputs set based on current step, not after condition evaluation
*)
(* CONTRACT_RULES [] *)

startRisingEdge(CLK := Start);

IF EmergencyStop = FALSE THEN
    MoveDown := FALSE;
    MoveUp := FALSE;
    MoveLeft := FALSE;
    MoveRight := FALSE;
    ActivateGrip := FALSE;
    ActivateRelease := FALSE;
    running := FALSE;
    cycleComplete := FALSE;
    step := 0;
ELSE
    IF ManualMode THEN
        step := 0;
        running := FALSE;
        MoveDown := DownButton AND NOT DownLimitSwitch;
        MoveUp := UpButton AND NOT UpLimitSwitch;
        MoveLeft := LeftButton AND NOT LeftLimitSwitch;
        MoveRight := RightButton AND NOT RightLimitSwitch;
        ActivateGrip := GripButton;
        ActivateRelease := ReleaseButton;

    ELSIF SingleStepMode THEN
        MoveDown := FALSE;
        MoveUp := FALSE;
        MoveLeft := FALSE;
        MoveRight := FALSE;
        ActivateGrip := FALSE;
        ActivateRelease := FALSE;

        IF startRisingEdge.Q AND NOT running THEN
            running := TRUE;
        END_IF;

        IF running THEN
            CASE step OF
                0:
                    IF NOT DownLimitSwitch THEN
                        MoveDown := TRUE;
                    END_IF;
                    IF DownLimitSwitch THEN
                        step := 1;
                        running := FALSE;
                    END_IF;
                1:
                    IF NOT GripLimitSwitch THEN
                        ActivateGrip := TRUE;
                    END_IF;
                    IF GripLimitSwitch THEN
                        step := 2;
                        running := FALSE;
                    END_IF;
                2:
                    IF NOT UpLimitSwitch THEN
                        MoveUp := TRUE;
                    END_IF;
                    IF UpLimitSwitch THEN
                        step := 3;
                        running := FALSE;
                    END_IF;
                3:
                    IF NOT RightLimitSwitch THEN
                        MoveRight := TRUE;
                    END_IF;
                    IF RightLimitSwitch THEN
                        step := 4;
                        running := FALSE;
                    END_IF;
                4:
                    IF NOT DownLimitSwitch THEN
                        MoveDown := TRUE;
                    END_IF;
                    IF DownLimitSwitch THEN
                        step := 5;
                        running := FALSE;
                    END_IF;
                5:
                    IF NOT ReleaseLimitSwitch THEN
                        ActivateRelease := TRUE;
                    END_IF;
                    IF ReleaseLimitSwitch THEN
                        step := 6;
                        running := FALSE;
                    END_IF;
                6:
                    IF NOT UpLimitSwitch THEN
                        MoveUp := TRUE;
                    END_IF;
                    IF UpLimitSwitch THEN
                        step := 7;
                        running := FALSE;
                    END_IF;
                7:
                    IF NOT LeftLimitSwitch THEN
                        MoveLeft := TRUE;
                    END_IF;
                    IF LeftLimitSwitch THEN
                        step := 0;
                        running := FALSE;
                    END_IF;
            END_CASE;
        END_IF;

    ELSIF SingleCycleMode THEN
        MoveDown := FALSE;
        MoveUp := FALSE;
        MoveLeft := FALSE;
        MoveRight := FALSE;
        ActivateGrip := FALSE;
        ActivateRelease := FALSE;

        IF startRisingEdge.Q AND NOT running AND NOT cycleComplete THEN
            running := TRUE;
        END_IF;

        IF running THEN
            CASE step OF
                0:
                    IF NOT DownLimitSwitch THEN
                        MoveDown := TRUE;
                    END_IF;
                    IF DownLimitSwitch THEN
                        step := 1;
                    END_IF;
                1:
                    IF NOT GripLimitSwitch THEN
                        ActivateGrip := TRUE;
                    END_IF;
                    IF GripLimitSwitch THEN
                        step := 2;
                    END_IF;
                2:
                    IF NOT UpLimitSwitch THEN
                        MoveUp := TRUE;
                    END_IF;
                    IF UpLimitSwitch THEN
                        step := 3;
                    END_IF;
                3:
                    IF NOT RightLimitSwitch THEN
                        MoveRight := TRUE;
                    END_IF;
                    IF RightLimitSwitch THEN
                        step := 4;
                    END_IF;
                4:
                    IF NOT DownLimitSwitch THEN
                        MoveDown := TRUE;
                    END_IF;
                    IF DownLimitSwitch THEN
                        step := 5;
                    END_IF;
                5:
                    IF NOT ReleaseLimitSwitch THEN
                        ActivateRelease := TRUE;
                    END_IF;
                    IF ReleaseLimitSwitch THEN
                        step := 6;
                    END_IF;
                6:
                    IF NOT UpLimitSwitch THEN
                        MoveUp := TRUE;
                    END_IF;
                    IF UpLimitSwitch THEN
                        step := 7;
                    END_IF;
                7:
                    IF NOT LeftLimitSwitch THEN
                        MoveLeft := TRUE;
                    END_IF;
                    IF LeftLimitSwitch THEN
                        running := FALSE;
                        cycleComplete := TRUE;
                        step := 0;
                    END_IF;
            END_CASE;
        END_IF;

    ELSIF ContinuousMode THEN
        MoveDown := FALSE;
        MoveUp := FALSE;
        MoveLeft := FALSE;
        MoveRight := FALSE;
        ActivateGrip := FALSE;
        ActivateRelease := FALSE;

        IF startRisingEdge.Q AND NOT running THEN
            running := TRUE;
        END_IF;

        IF running THEN
            CASE step OF
                0:
                    IF NOT DownLimitSwitch THEN
                        MoveDown := TRUE;
                    END_IF;
                    IF DownLimitSwitch THEN
                        step := 1;
                    END_IF;
                1:
                    IF NOT GripLimitSwitch THEN
                        ActivateGrip := TRUE;
                    END_IF;
                    IF GripLimitSwitch THEN
                        step := 2;
                    END_IF;
                2:
                    IF NOT UpLimitSwitch THEN
                        MoveUp := TRUE;
                    END_IF;
                    IF UpLimitSwitch THEN
                        step := 3;
                    END_IF;
                3:
                    IF NOT RightLimitSwitch THEN
                        MoveRight := TRUE;
                    END_IF;
                    IF RightLimitSwitch THEN
                        step := 4;
                    END_IF;
                4:
                    IF NOT DownLimitSwitch THEN
                        MoveDown := TRUE;
                    END_IF;
                    IF DownLimitSwitch THEN
                        step := 5;
                    END_IF;
                5:
                    IF NOT ReleaseLimitSwitch THEN
                        ActivateRelease := TRUE;
                    END_IF;
                    IF ReleaseLimitSwitch THEN
                        step := 6;
                    END_IF;
                6:
                    IF NOT UpLimitSwitch THEN
                        MoveUp := TRUE;
                    END_IF;
                    IF UpLimitSwitch THEN
                        step := 7;
                    END_IF;
                7:
                    IF NOT LeftLimitSwitch THEN
                        MoveLeft := TRUE;
                    END_IF;
                    IF LeftLimitSwitch THEN
                        step := 0;
                    END_IF;
            END_CASE;
        END_IF;
    END_IF;
END_IF;

END_FUNCTION_BLOCK

(* ---- public-hard-06.candidate_01.st ---- *)
(* ENGINEERING_CONTRACT *)
(*
┌──────────────────┬────────────────────────────────────────────────────────────────────────┐
│ Output/State     │ Activation, Retention, Reset, Priority, Units                          │
├──────────────────┼────────────────────────────────────────────────────────────────────────┤
│ MotorForward     │ Active during FEED, TRANSPORT_TO_WEIGH, TRANSPORT_TO_FIRING states     │
│                  │ in automatic mode only. Deactivated on state exit. PUB003, PUB006      │
├──────────────────┼────────────────────────────────────────────────────────────────────────┤
│ MotorReverse     │ Active during KICK state only (automatic mode). Deactivated on exit.   │
│                  │ Interlocked with MotorForward in manual mode. PUB002                   │
├──────────────────┼────────────────────────────────────────────────────────────────────────┤
│ kick             │ Latched HIGH when weight < 100 OR weight > 200 in WEIGH state.         │
│                  │ Deactivated when material exits wash station (SensorWash=FALSE).       │
│                  │ Single rejection per material cycle. PUB010                            │
├──────────────────┼────────────────────────────────────────────────────────────────────────┤
│ CompletionLight  │ Latched HIGH when SensorOutput=TRUE in OUTPUT state.                   │
│                  │ Deactivated when SensorOutput=FALSE (product removed).                 │
│                  │ No manual override specified. PUB012                                   │
├──────────────────┼────────────────────────────────────────────────────────────────────────┤
│ firingTemp       │ Calculated once when weight passes qualification check.                │
│                  │ Value: 500 + (weight - 100) * 0.5, range [500, 550]. Retained.         │
│                  │ PUB011                                                                   │
├──────────────────┼────────────────────────────────────────────────────────────────────────┤
│ State Machine    │ States: IDLE(0), FEED(1), WASH_WAIT(2), WEIGH(3), KICK(4),             │
│                  │ TRANSPORT_TO_FIRING(5), FIRING_WAIT(6), TRANSPORT_TO_OUTPUT(7),        │
│                  │ OUTPUT(8). Same-scan priority: sensor arrival > state transition.      │
│                  │ PUB003-PUB012                                                           │
└──────────────────┴────────────────────────────────────────────────────────────────────────┘
*)

(* CONTRACT_RULES [{"kind":"hold_until_reset","output":"CompletionLight","set_input":"SensorOutput","reset_input":"NOT SensorOutput"}] *)

FUNCTION_BLOCK ProductionControl
VAR
    tmp_state : INT := 0;
    tmp_prevSensorFeed : BOOL := FALSE;
    tmp_prevSensorWash : BOOL := FALSE;
    tmp_prevSensorWeight : BOOL := FALSE;
    tmp_prevSensorFiring : BOOL := FALSE;
END_VAR

// Reset all outputs at start of scan
MotorForward := FALSE;
MotorReverse := FALSE;
kick := FALSE;
CompletionLight := FALSE;

IF Mode = FALSE THEN
    // Manual Mode (PUB001, PUB002)
    MotorForward := ForwardButton AND NOT ReverseButton;
    MotorReverse := ReverseButton AND NOT ForwardButton;
ELSE
    // Automatic Mode (PUB003-PUB012)
    CASE tmp_state OF
        0: // IDLE - waiting for material at feed station
            IF SensorFeed THEN
                tmp_state := 1;
            END_IF;

        1: // FEED - transport to cleaning station
            MotorForward := TRUE;
            IF SensorWash THEN
                tmp_state := 2;
                MotorForward := FALSE;
            END_IF;

        2: // WASH_WAIT - waiting for cleaning completion
            IF washComplete THEN
                tmp_state := 3;
            END_IF;

        3: // WEIGH - process weight measurement
            IF weightComplete THEN
                IF weight < 100.0 OR weight > 200.0 THEN
                    // Unqualified: initiate kick
                    kick := TRUE;
                    MotorReverse := TRUE;
                    tmp_state := 4;
                ELSE
                    // Qualified: calculate firing temperature
                    firingTemp := 500.0 + (weight - 100.0) * 0.5;
                    MotorForward := TRUE;
                    tmp_state := 5;
                END_IF;
            END_IF;

        4: // KICK - reverse transport to exit wash station
            kick := TRUE;
            MotorReverse := TRUE;
            IF NOT SensorWash THEN
                kick := FALSE;
                MotorReverse := FALSE;
                tmp_state := 0;
            END_IF;

        5: // TRANSPORT_TO_FIRING
            MotorForward := TRUE;
            IF SensorFiring THEN
                tmp_state := 6;
                MotorForward := FALSE;
            END_IF;

        6: // FIRING_WAIT - waiting for firing completion
            IF firingComplete THEN
                tmp_state := 7;
            END_IF;

        7: // TRANSPORT_TO_OUTPUT
            MotorForward := TRUE;
            IF SensorOutput THEN
                tmp_state := 8;
                MotorForward := FALSE;
            END_IF;

        8: // OUTPUT - product complete, light on
            IF SensorOutput THEN
                CompletionLight := TRUE;
            ELSE
                CompletionLight := FALSE;
                tmp_state := 0;
            END_IF;

    END_CASE;
END_IF;

END_FUNCTION_BLOCK

(* ---- public-hard-06.candidate_02.st ---- *)
(* ENGINEERING_CONTRACT *)
(*
┌──────────────────┬────────────────────────────────────────────────────────────────────────┐
│ Output/State     │ Activation, Retention, Reset, Priority, Units                          │
├──────────────────┼────────────────────────────────────────────────────────────────────────┤
│ MotorForward     │ Active during FEED, TRANSPORT_TO_WEIGH, TRANSPORT_TO_FIRING states     │
│                  │ in automatic mode only. Deactivated on state exit. PUB003, PUB006      │
├──────────────────┼────────────────────────────────────────────────────────────────────────┤
│ MotorReverse     │ Active during KICK state only (automatic mode). Deactivated on exit.   │
│                  │ Interlocked with MotorForward in manual mode. PUB002                   │
├──────────────────┼────────────────────────────────────────────────────────────────────────┤
│ kick             │ Latched HIGH when weight < 100 OR weight > 200 in WEIGH state.         │
│                  │ Deactivated when material exits wash station (SensorWash=FALSE).       │
│                  │ Single rejection per material cycle. PUB010                            │
├──────────────────┼────────────────────────────────────────────────────────────────────────┤
│ CompletionLight  │ Latched HIGH when SensorOutput=TRUE in OUTPUT state.                   │
│                  │ Deactivated when SensorOutput=FALSE (product removed).                 │
│                  │ No manual override specified. PUB012                                   │
├──────────────────┼────────────────────────────────────────────────────────────────────────┤
│ firingTemp       │ Calculated once when weight passes qualification check.                │
│                  │ Value: 500 + (weight - 100) * 0.5, range [500, 550]. Retained.         │
│                  │ PUB011                                                                   │
├──────────────────┼────────────────────────────────────────────────────────────────────────┤
│ State Machine    │ States: IDLE(0), FEED(1), WASH_WAIT(2), WEIGH(3), KICK(4),             │
│                  │ TRANSPORT_TO_FIRING(5), FIRING_WAIT(6), TRANSPORT_TO_OUTPUT(7),        │
│                  │ OUTPUT(8). Same-scan priority: sensor arrival > state transition.      │
│                  │ PUB003-PUB012                                                           │
└──────────────────┴────────────────────────────────────────────────────────────────────────┘
*)

(* CONTRACT_RULES [{"kind":"hold_until_reset","output":"CompletionLight","set_input":"SensorOutput","reset_input":"NOT SensorOutput"}] *)

FUNCTION_BLOCK ProductionControl
VAR_INPUT
    Mode : BOOL;
    ForwardButton : BOOL;
    ReverseButton : BOOL;
    SensorFeed : BOOL;
    SensorWash : BOOL;
    SensorWeight : BOOL;
    SensorFiring : BOOL;
    SensorOutput : BOOL;
    washComplete : BOOL;
    weightComplete : BOOL;
    weight : REAL;
    firingComplete : BOOL;
END_VAR

VAR_OUTPUT
    MotorForward : BOOL;
    MotorReverse : BOOL;
    kick : BOOL;
    CompletionLight : BOOL;
    firingTemp : REAL;
END_VAR

VAR
    tmp_state : INT := 0;
    tmp_prevSensorFeed : BOOL := FALSE;
    tmp_prevSensorWash : BOOL := FALSE;
    tmp_prevSensorWeight : BOOL := FALSE;
    tmp_prevSensorFiring : BOOL := FALSE;
END_VAR

// Reset all outputs at start of scan
MotorForward := FALSE;
MotorReverse := FALSE;
kick := FALSE;
CompletionLight := FALSE;

IF Mode = FALSE THEN
    // Manual Mode (PUB001, PUB002)
    MotorForward := ForwardButton AND NOT ReverseButton;
    MotorReverse := ReverseButton AND NOT ForwardButton;
ELSE
    // Automatic Mode (PUB003-PUB012)
    CASE tmp_state OF
        0: // IDLE - waiting for material at feed station
            IF SensorFeed THEN
                tmp_state := 1;
            END_IF;

        1: // FEED - transport to cleaning station
            MotorForward := TRUE;
            IF SensorWash THEN
                tmp_state := 2;
                MotorForward := FALSE;
            END_IF;

        2: // WASH_WAIT - waiting for cleaning completion
            IF washComplete THEN
                tmp_state := 3;
            END_IF;

        3: // WEIGH - process weight measurement
            IF weightComplete THEN
                IF weight < 100.0 OR weight > 200.0 THEN
                    // Unqualified: initiate kick
                    kick := TRUE;
                    MotorReverse := TRUE;
                    tmp_state := 4;
                ELSE
                    // Qualified: calculate firing temperature
                    firingTemp := 500.0 + (weight - 100.0) * 0.5;
                    MotorForward := TRUE;
                    tmp_state := 5;
                END_IF;
            END_IF;

        4: // KICK - reverse transport to exit wash station
            kick := TRUE;
            MotorReverse := TRUE;
            IF NOT SensorWash THEN
                kick := FALSE;
                MotorReverse := FALSE;
                tmp_state := 0;
            END_IF;

        5: // TRANSPORT_TO_FIRING
            MotorForward := TRUE;
            IF SensorFiring THEN
                tmp_state := 6;
                MotorForward := FALSE;
            END_IF;

        6: // FIRING_WAIT - waiting for firing completion
            IF firingComplete THEN
                tmp_state := 7;
            END_IF;

        7: // TRANSPORT_TO_OUTPUT
            MotorForward := TRUE;
            IF SensorOutput THEN
                tmp_state := 8;
                MotorForward := FALSE;
            END_IF;

        8: // OUTPUT - product complete, light on
            IF SensorOutput THEN
                CompletionLight := TRUE;
            ELSE
                CompletionLight := FALSE;
                tmp_state := 0;
            END_IF;

    END_CASE;
END_IF;

END_FUNCTION_BLOCK

(* ---- public-hard-06.candidate_03.st ---- *)
(* ENGINEERING_CONTRACT *)
(*
┌──────────────────┬────────────────────────────────────────────────────────────────────────┐
│ Output/State     │ Activation, Retention, Reset, Priority, Units                          │
├──────────────────┼────────────────────────────────────────────────────────────────────────┤
│ MotorForward     │ Active during FEED, TRANSPORT_TO_WEIGH, TRANSPORT_TO_FIRING states     │
│                  │ in automatic mode only. Deactivated on state exit. PUB003, PUB006      │
├──────────────────┼────────────────────────────────────────────────────────────────────────┤
│ MotorReverse     │ Active during KICK state only (automatic mode). Deactivated on exit.   │
│                  │ Interlocked with MotorForward in manual mode. PUB002                   │
├──────────────────┼────────────────────────────────────────────────────────────────────────┤
│ kick             │ Latched HIGH when weight < 100 OR weight > 200 in WEIGH state.         │
│                  │ Deactivated when material exits wash station (SensorWash=FALSE).       │
│                  │ Single rejection per material cycle. PUB010                            │
├──────────────────┼────────────────────────────────────────────────────────────────────────┤
│ CompletionLight  │ Latched HIGH when SensorOutput=TRUE in OUTPUT state.                   │
│                  │ Deactivated when SensorOutput=FALSE (product removed).                 │
│                  │ No manual override specified. PUB012                                   │
├──────────────────┼────────────────────────────────────────────────────────────────────────┤
│ firingTemp       │ Calculated once when weight passes qualification check.                │
│                  │ Value: 500 + (weight - 100) * 0.5, range [500, 550]. Retained.         │
│                  │ PUB011                                                                   │
├──────────────────┼────────────────────────────────────────────────────────────────────────┤
│ State Machine    │ States: IDLE(0), FEED(1), WASH_WAIT(2), WEIGH(3), KICK(4),             │
│                  │ TRANSPORT_TO_FIRING(5), FIRING_WAIT(6), TRANSPORT_TO_OUTPUT(7),        │
│                  │ OUTPUT(8). Same-scan priority: sensor arrival > state transition.      │
│                  │ PUB003-PUB012                                                           │
└──────────────────┴────────────────────────────────────────────────────────────────────────┘
*)

(* CONTRACT_RULES [{"kind":"hold_until_reset","output":"CompletionLight","set_input":"SensorOutput","reset_input":"NOT SensorOutput"}] *)

FUNCTION_BLOCK ProductionControl
VAR_INPUT
    Mode : BOOL;
    ForwardButton : BOOL;
    ReverseButton : BOOL;
    SensorFeed : BOOL;
    SensorWash : BOOL;
    SensorWeight : BOOL;
    SensorFiring : BOOL;
    SensorOutput : BOOL;
    washComplete : BOOL;
    weightComplete : BOOL;
    weight : REAL;
    firingComplete : BOOL;
END_VAR

VAR_OUTPUT
    MotorForward : BOOL;
    MotorReverse : BOOL;
    kick : BOOL;
    CompletionLight : BOOL;
    firingTemp : REAL;
END_VAR

VAR
    tmp_state : INT := 0;
END_VAR

// Reset all outputs at start of scan
MotorForward := FALSE;
MotorReverse := FALSE;
kick := FALSE;
CompletionLight := FALSE;

IF Mode = FALSE THEN
    // Manual Mode (PUB001, PUB002)
    MotorForward := ForwardButton AND NOT ReverseButton;
    MotorReverse := ReverseButton AND NOT ForwardButton;
ELSE
    // Automatic Mode (PUB003-PUB012)
    CASE tmp_state OF
        0: // IDLE - waiting for material at feed station
            IF SensorFeed THEN
                tmp_state := 1;
                MotorForward := TRUE;
            END_IF;

        1: // FEED - transport to cleaning station
            MotorForward := TRUE;
            IF SensorWash THEN
                tmp_state := 2;
                MotorForward := FALSE;
            END_IF;

        2: // WASH_WAIT - waiting for cleaning completion
            IF washComplete THEN
                tmp_state := 3;
            END_IF;

        3: // WEIGH - process weight measurement
            IF weightComplete THEN
                IF weight < 100.0 OR weight > 200.0 THEN
                    // Unqualified: initiate kick
                    kick := TRUE;
                    MotorReverse := TRUE;
                    tmp_state := 4;
                ELSE
                    // Qualified: calculate firing temperature
                    firingTemp := 500.0 + (weight - 100.0) * 0.5;
                    MotorForward := TRUE;
                    tmp_state := 5;
                END_IF;
            END_IF;

        4: // KICK - reverse transport to exit wash station
            kick := TRUE;
            MotorReverse := TRUE;
            IF NOT SensorWash THEN
                kick := FALSE;
                MotorReverse := FALSE;
                tmp_state := 0;
            END_IF;

        5: // TRANSPORT_TO_FIRING
            MotorForward := TRUE;
            IF SensorFiring THEN
                tmp_state := 6;
                MotorForward := FALSE;
            END_IF;

        6: // FIRING_WAIT - waiting for firing completion
            IF firingComplete THEN
                tmp_state := 7;
            END_IF;

        7: // TRANSPORT_TO_OUTPUT
            MotorForward := TRUE;
            IF SensorOutput THEN
                tmp_state := 8;
                MotorForward := FALSE;
            END_IF;

        8: // OUTPUT - product complete, light on
            IF SensorOutput THEN
                CompletionLight := TRUE;
            ELSE
                CompletionLight := FALSE;
                tmp_state := 0;
            END_IF;

    END_CASE;
END_IF;

END_FUNCTION_BLOCK
